Yaskawa INFORM job: TGTPROG.JBI

/JOB
//NAME TGTPROG
//POS
///NPOS 2,0,0,0,0,0
///TOOL 9
///POSTYPE PULSE
///PULSE
C00000=10240,-20480,45966,-57458,68949,-40619,34475
C00001=512,-256,-1724,3160,-3519,580,144
//INST
<volatile>
///COMM Generated using RoboDK
///ATTR SC,RW
///GROUP1 RB1
NOP
'Program generated by RoboDK v
'6.0.7 for Yaskawa Motoman SIA
' on XX/XX/XXXX 18:00:00
'Using nominal kinematics.
MOVJ C00000 VJ=50.00
MOVL C00001 V=100.0
END
